// TIA Portal V21 export
VAR_GLOBAL   // PLC tag table "ModeConstant"
END_VAR
VAR_GLOBAL CONSTANT   // user constants
   PLACE_LOCAL : Int := 3;
   PLACE_PU1 : Int := 0;
   PLACE_PU2 : Int := 1;
   PLACE_DISPATCHER : Int := 2;
   MODE_SERVICE : Int := 1;
   MODE_SEMIAUTO : Int := 4;
   MODE_DISABLE : Int := 0;
   MODE_AUTO : Int := 8;
   MODE_MANUAL : Int := 2;
END_VAR
